// TIA Portal V21 export
// export: Created 2026-10-23T20:42:23.8551304Z, ExportSetting WithDefaults, DisplayName Totally Integrated Automation Portal, DisplayVersion V21 Update 1, DisplayName SINAMICS Startdrive Advanced, DisplayVersion V21 HF2, DisplayName SINAMICS Startdrive G110M, G120, G120C, G120D, G120P, G115D, DisplayVersion V21 HF2, DisplayName SINAMICS Startdrive G130, G150, S120, S150, G200, G220, S200, S210, S220, Innomotics MVD, DisplayVersion V21 HF2, DisplayName STEP 7 Professional, DisplayVersion V21 Update 1, DisplayName STEP 7 Safety, DisplayVersion V21, DisplayName Tech WebApplication, DisplayVersion V21, DisplayName WinCC Basic/Comfort/Advanced, DisplayVersion V21 Update 1, DisplayName WinCC Unified, DisplayVersion V21 Update 1
FUNCTION_BLOCK "FB_SclTimers"   // FB2, SCL
TITLE = IEC timers, counters and edges
{ S7_Optimized_Access := 'TRUE' }
VERSION : 0.1
// Every IEC timer, edge and counter as a multi-instance, each called every cycle
// stored: AutoNumber true, IsIECCheckEnabled false, IsRetainMemResEnabled false, MemoryReserve 100, SetENOAutomatically false, UDAEnableTagReadback false
   VAR_INPUT
      Start : Bool;   // Start signal
      Reset : Bool;   // Reset the counter
      DelayTime : Time := T#2S;   // On-delay time
   END_VAR
   VAR_OUTPUT
      DelayedOn : Bool;   // Start delayed by DelayTime
      RunOn : Bool;   // Start with run-on time
      Pulse : Bool;   // Pulse on the rising edge of Start
      Count : Int;   // Number of falling edges of Start
      CountReached : Bool;   // Count has reached the preset
   END_VAR
   VAR
      OnDelay { S7_SetPoint := 'True'} : TON_TIME;   // On-delay timer
      OffDelay { S7_SetPoint := 'True'} : TOF_TIME;   // Off-delay timer
      PulseTimer { S7_SetPoint := 'True'} : TP_TIME;   // Pulse timer
      StartEdge { S7_SetPoint := 'True'} : R_TRIG;   // Rising edge of Start
      StopEdge { S7_SetPoint := 'True'} : F_TRIG;   // Falling edge of Start
      PartCounter { S7_SetPoint := 'True'} : CTU_INT;   // Up counter
   END_VAR
   VAR CONSTANT
      COUNT_PRESET : Int := 10;   // Counter preset
   END_VAR
BEGIN

       REGION Timers
           #OnDelay(IN := #Start, PT := #DelayTime, Q => #DelayedOn);
           #OffDelay(IN := #Start, PT := T#3s, Q => #RunOn);
       END_REGION

       REGION Edges and pulse
           #StartEdge(CLK := #Start);
           #StopEdge(CLK := #Start);
           #PulseTimer(IN := #StartEdge.Q, PT := T#500ms, Q => #Pulse);
       END_REGION

       REGION Counter
           #PartCounter(CU := #StopEdge.Q, R := #Reset, PV := #COUNT_PRESET, Q => #CountReached, CV => #Count);
       END_REGION
END_FUNCTION_BLOCK
